(* IEC 61131-3 sources: codesys-framework/txt/application/WeVe IO (library)/Analog Input, 5 files *)

(* ---- E_AnalogInputType.dut.st ---- *)
TYPE E_AnalogInputType :
(
	Invalid := 0,
	S401_0_10V := 1,
	S401_1_5V := 2
);
END_TYPE

(* ---- E_EngineeringUnits.dut.st ---- *)
TYPE E_EngineeringUnits :
(
	Volt := 0,
	gram := 1,
	bar :=2,
	degree :=3,
	cubicmeters :=4,
	milimeters := 5,
	G := 6
);
END_TYPE

(* ---- SC_AnalogInputSignals.dut.st ---- *)
TYPE SC_AnalogInputSignals :
STRUCT
	iRawValue 	: INT;
	rValue 		: REAL;
	sUnit 		: STRING (20);
END_STRUCT
END_TYPE

(* ---- SC_SystemParametersAnalogInput.dut.st ---- *)
TYPE SC_SystemParametersAnalogInput :
STRUCT
	eAI_Type	 							: E_AnalogInputType;
	eSignalEngUnit 							: E_EngineeringUnits;
	rSignalValueEngUnit_AnalogMinLevel 		: REAL;
	rSignalValueEngUnit_AnalogMaxLevel 		: REAL;
	rSignalValueEngUnit_atAnalogMinLevel 	: REAL;
	rSignalValueEngUnit_atAnalogMaxLevel 	: REAL;
END_STRUCT
END_TYPE

(* ---- FB_AnalogInput.pou.st ---- *)
FUNCTION_BLOCK FB_AnalogInput
VAR_INPUT
	iAI_Value 		: INT;
END_VAR
VAR_OUTPUT
END_VAR
VAR
	_scSysPar 			: SC_SystemParametersAnalogInput;
	_scSignalValue 		: SC_AnalogInputSignals;
END_VAR

// --- BEGIN IMPLEMENTATION ---

// Scale output value (dependant on input signal type)
_scSignalValue.iRawValue := iAI_Value;

_scSignalValue.rValue := F_Scale (
	rInputScaleValue := INT_TO_REAL(iAI_Value),
	rInputScaleValueMinLevel := _scSysPar.rSignalValueEngUnit_AnalogMinLevel,
	rInputScaleValueMaxLevel := _scSysPar.rSignalValueEngUnit_AnalogMaxLevel,
	rOutputScaleValueMinLevel := _scSysPar.rSignalValueEngUnit_atAnalogMinLevel,
	rOutputScaleValueMaxLevel := _scSysPar.rSignalValueEngUnit_atAnalogMaxLevel,
	eScaleMethod := E_ScaleMethod.ExtraPolation);

// Add EngineeringUnitString
_scSignalValue.sUnit := F_GetEngUnit(_scSysPar.eSignalEngUnit);
